(* IEC 61131-3 sources: kns-port-domestic/tools/inventory_tests/fixtures/lib/src/POUs/FB_Child, 1 file *)

(* ---- FB_Child.decl.st ---- *)
// Назначение: наследник базы
FUNCTION_BLOCK FINAL FB_Child EXTENDS FB_Base
VAR_IN_OUT
    stExt : ST_Ext;
END_VAR
